{attribute 'qualified_only'}
VAR_GLOBAL
  bQrEnabled     : BOOL := FALSE;
  bQrCodeFound   : BOOL := FALSE;
  bQrCameraConnected : BOOL := FALSE; // Camera hardware connected
  bQrActive      : BOOL := FALSE;    // Enabled OR camera connected (VISU lamp)
  sQrCodeText    : STRING(255) := '';
  sQrDisplayText : STRING(512) := 'QR scanner OFF';
  hrQrVision     : HRESULT := 0;
END_VAR

(* stored: Version 1.1.0.1, ProductVersion 3.1.4026.17
   GVL GVL_Data: Id {e207c451-feb9-482c-923f-2b3efa1bd73d} *)
